// Mitsubishi GX Works2 project: 261012_타이머실습_클럭펄스   PLC: Q03UDV

PROGRAM MAIN
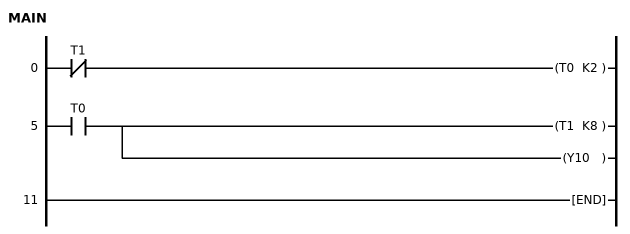
0     LDI     T1
      OUT     T0 K2
5     LD      T0
      OUT     T1 K8
      OUT     Y10
11    END
END_PROGRAM
